Staubli VAL3: onStart.pgx

program onStart()
  local num l_nSize
  local num l_i
begin
  l_nSize=size(savedata:fFrameItem)
  resize(sFrameList,1,l_nSize)
  l_nSize=size(savedata:tToolItem)
  resize(sToolList,1,l_nSize)

  for l_i = 0 to size(sFrameList)-1
    sFrameList[l_i]=toString("",l_i)+","+savedata:fFrameItem[l_i].sName
  endFor

  for l_i = 0 to size(sToolList)-1
    sToolList[l_i]=toString("",l_i)+","+savedata:tToolItem[l_i].sName
  endFor

  sSelFrame=sFrameList[0]
  sSelTool=sToolList[0]

end
